// TIA Portal V20 export
// export: Created 2026-10-21T13:28:38.0844279Z, ExportSetting None, DisplayName Totally Integrated Automation Portal, DisplayVersion V20, DisplayName TIA Portal Openness, DisplayVersion V20, DisplayName TIA Portal Version Control Interface, DisplayVersion V20, DisplayName STEP 7 Professional, DisplayVersion V20, DisplayName STEP 7 Safety, DisplayVersion V20, DisplayName WinCC Basic/Comfort/Advanced, DisplayVersion V20, DisplayName WinCC Unified, DisplayVersion V20
VAR_GLOBAL   // PLC tag table "Cinta_Signals"
   DI_ES01_Ok AT %M0.0 : Bool;
   DI_M01_Start AT %M0.1 : Bool;
   DI_M01_Stop AT %M0.2 : Bool;
   DI_M01_Reset AT %M0.3 : Bool;
   DI_M01_Feedback AT %M0.4 : Bool;
   DO_M01_Run AT %M1.0 : Bool;
   M_M01_Running AT %M1.1 : Bool;
   M_M01_Interlock AT %M1.2 : Bool;
   M_M01_Fault AT %M1.3 : Bool;
   M_M01_FaultCode AT %MW4 : Int;
END_VAR
